Fanuc KAREL source: kc00021.KL

-- PROVISIONAL review KL for V1013-1; original PC SHA256 edc3aaf1c179a914ec167f89cecd04b1683a33f1c04ccd45abad6b92ab5ac89a
-- Incomplete behavior may be omitted. Consult companion uncertainty JSON. Do not deploy.
PROGRAM KC00021
%NOLOCKGROUP
BEGIN
  -- UNRESOLVED_PC offsets 5-18; opcodes 27,27,27,9C,31,23
  -- UNRESOLVED_PC offsets 23-27; opcodes 7F
END KC00021
